Fanuc KAREL source: KB00043.KL

PROGRAM KB00043
%NOLOCKGROUP
%ENVIRONMENT TIM
VAR
  P1: INTEGER
  P2: STRING[80]
BEGIN
  P1 = 1
  P2 = 'A'
  CNV_TIME_STR(P1, P2)
END KB00043
